FUNCTION_BLOCK FB_Line_Target EXTENDS FB_SFC_Cycle IMPLEMENTS ITF_FB_SFC_Cycle
VAR_INPUT
	valTankA				:	E_Pis_Name	;
	valTankB				:	E_Pis_Name	;
	valTankA_Pipe			:	E_Pis_Name	;
	valTankB_Pipe			:	E_Pis_Name	;
	valDrain				:	E_Pis_Name	;
	valCIP					:	E_Pis_Name	;
END_VAR
VAR_OUTPUT
END_VAR
VAR
	eReq				: E_Line_Target;
	eProcess			: E_Line_Target;
	eStatus				: E_Line_Target;
	
	fbPis				: FB_Piston;
	
	stPis_TankA				: REFERENCE TO ST_Piston;
	stPis_TankB				: REFERENCE TO ST_Piston;
	stPis_TankA_Pipe		: REFERENCE TO ST_Piston;
	stPis_TankB_Pipe		: REFERENCE TO ST_Piston;
	stPis_Drain				: REFERENCE TO ST_Piston;
	stPis_CIP				: REFERENCE TO ST_Piston;
	
	stPis_Outlet: ST_Piston;
	tonDrainTime: TON;
	rt_Req_Reset: R_TRIG;
END_VAR

act_GetReference();

act_Oper();
//IF NOT Init.x THEN
	act_Status();
//END_IF

tonDrainTime(PT:=T#1M, IN:=eStatus=E_Line_Target.eDrain AND eReq=E_Line_Target.eNone);
IF tonDrainTime.Q 
AND eReq=E_Line_Target.eNone
AND eProcess=E_Line_Target.eNone
THEN;
	eReq:=E_Line_Target.eClose;
END_IF

m_Request_Reset(memo:=rt_Req_Reset);//

ACTION _aCIP_active:
bStepDone:=FALSE;
IF TRUE 
AND eStatus=E_Line_Target.eCIP
THEN;
	bStepDone:=TRUE;
END_IF
END_ACTION

ACTION _aCIP_entry:
fbPis.m_SetByRecipe(stPis:=stPis_TankA, 			req:=E_Piston_Recipe_State.Release);
//fbPis.m_SetByRecipe(stPis:=stPis_TankA_Pipe, 		req:=E_Piston_Recipe_State.Release);		
fbPis.m_SetByRecipe(stPis:=stPis_TankB, 			req:=E_Piston_Recipe_State.Release);
//fbPis.m_SetByRecipe(stPis:=stPis_TankB_Pipe, 		req:=E_Piston_Recipe_State.Release);
fbPis.m_SetByRecipe(stPis:=stPis_Drain, 			req:=E_Piston_Recipe_State.Act);
fbPis.m_SetByRecipe(stPis:=stPis_CIP, 				req:=E_Piston_Recipe_State.Act);
END_ACTION

ACTION _aClose_active:
bStepDone:=FALSE;
IF TRUE 
AND eStatus=E_Line_Target.eClose
THEN;
	bStepDone:=TRUE;
END_IF
END_ACTION

ACTION _aClose_entry:
fbPis.m_SetByRecipe(stPis:=stPis_TankA, 			req:=E_Piston_Recipe_State.Release);
//fbPis.m_SetByRecipe(stPis:=stPis_TankA_Pipe, 		req:=E_Piston_Recipe_State.Release);		
fbPis.m_SetByRecipe(stPis:=stPis_TankB, 			req:=E_Piston_Recipe_State.Release);
//fbPis.m_SetByRecipe(stPis:=stPis_TankB_Pipe, 		req:=E_Piston_Recipe_State.Release);
fbPis.m_SetByRecipe(stPis:=stPis_Drain, 			req:=E_Piston_Recipe_State.Release);
fbPis.m_SetByRecipe(stPis:=stPis_CIP, 				req:=E_Piston_Recipe_State.Release);
END_ACTION

ACTION _aDone_entry:
eProcess:=E_Line_Target.eNone;
eReq:=E_Line_Target.eNone;
bRun:=FALSE;
bDone:=TRUE;
END_ACTION

ACTION _aDrain_active:
bStepDone:=FALSE;
IF TRUE 
AND eStatus=E_Line_Target.eDrain
THEN;
	bStepDone:=TRUE;
END_IF
END_ACTION

ACTION _aDrain_entry:
fbPis.m_SetByRecipe(stPis:=stPis_TankA, 			req:=E_Piston_Recipe_State.Release);	
//fbPis.m_SetByRecipe(stPis:=stPis_TankA_Pipe, 		req:=E_Piston_Recipe_State.Release);	
fbPis.m_SetByRecipe(stPis:=stPis_TankB, 			req:=E_Piston_Recipe_State.Release);
//fbPis.m_SetByRecipe(stPis:=stPis_TankB_Pipe, 		req:=E_Piston_Recipe_State.Release);
fbPis.m_SetByRecipe(stPis:=stPis_Drain, 			req:=E_Piston_Recipe_State.Act);
fbPis.m_SetByRecipe(stPis:=stPis_CIP, 				req:=E_Piston_Recipe_State.Release);
END_ACTION

ACTION _aInit_active:
SFCReset:=FALSE;
END_ACTION

ACTION _aInit_exit:
eProcess:=E_Line_Target.eNone;
eReq:=E_Line_Target.eNone;
END_ACTION

ACTION _aReady_active:
CASE eReq OF
	E_Line_Target.eClose:;
			IF TRUE THEN;
				eProcess:=E_Line_Target.eClose;
			END_IF

	E_Line_Target.eTank_A:;
			IF TRUE THEN;
				eProcess:=E_Line_Target.eTank_A;
			END_IF	
			
	E_Line_Target.eTank_B:;
			IF TRUE THEN;
				eProcess:=E_Line_Target.eTank_B;
			END_IF	
			
	E_Line_Target.eCIP:;
			IF TRUE THEN;
				eProcess:=E_Line_Target.eCIP;
			END_IF	

	E_Line_Target.eDrain:;
			IF TRUE THEN;
				eProcess:=E_Line_Target.eDrain;
			END_IF	
		
END_CASE
END_ACTION

ACTION _aReady_exit:
bRun:=TRUE;
bDone:=FALSE;
END_ACTION

ACTION _aTank_A_active:
bStepDone:=FALSE;
IF TRUE  
AND eStatus=E_Line_Target.eTank_A 
THEN;
	bStepDone:=TRUE;
END_IF
END_ACTION

ACTION _aTank_A_entry:
fbPis.m_SetByRecipe(stPis:=stPis_TankA, 			req:=E_Piston_Recipe_State.Act);	
fbPis.m_SetByRecipe(stPis:=stPis_TankA_Pipe, 		req:=E_Piston_Recipe_State.Release);	
fbPis.m_SetByRecipe(stPis:=stPis_TankB, 			req:=E_Piston_Recipe_State.Release);
//fbPis.m_SetByRecipe(stPis:=stPis_TankB_Pipe, 		req:=E_Piston_Recipe_State.Release);
fbPis.m_SetByRecipe(stPis:=stPis_Drain, 			req:=E_Piston_Recipe_State.Release);
fbPis.m_SetByRecipe(stPis:=stPis_CIP, 				req:=E_Piston_Recipe_State.Release);
END_ACTION

ACTION _aTank_B_active:
bStepDone:=FALSE;
IF TRUE 
AND eStatus=E_Line_Target.eTank_B
THEN;
	bStepDone:=TRUE;
END_IF
END_ACTION

ACTION _aTank_B_entry:
fbPis.m_SetByRecipe(stPis:=stPis_TankA, 			req:=E_Piston_Recipe_State.Release);	
//fbPis.m_SetByRecipe(stPis:=stPis_TankA_Pipe, 		req:=E_Piston_Recipe_State.Release);	
fbPis.m_SetByRecipe(stPis:=stPis_TankB, 			req:=E_Piston_Recipe_State.Act);
fbPis.m_SetByRecipe(stPis:=stPis_TankB_Pipe, 		req:=E_Piston_Recipe_State.Release);
fbPis.m_SetByRecipe(stPis:=stPis_Drain, 			req:=E_Piston_Recipe_State.Release);
fbPis.m_SetByRecipe(stPis:=stPis_CIP, 				req:=E_Piston_Recipe_State.Release);
END_ACTION

ACTION act_GetReference:
m_Set_SFCFlags_Reference();
//refElement REF= fbElement[eElementID];
//refState_Long REF= fbElement[eElementID].eState_Long;

stPis_TankA				REF= g_Piston.stPis[valTankA];
stPis_TankB				REF= g_Piston.stPis[valTankB];
stPis_TankA_Pipe		REF= g_Piston.stPis[valTankA_Pipe];
stPis_TankB_Pipe		REF= g_Piston.stPis[valTankB_Pipe];
stPis_Drain				REF= g_Piston.stPis[valDrain];
stPis_CIP				REF= g_Piston.stPis[valCIP];
END_ACTION

ACTION act_Oper:
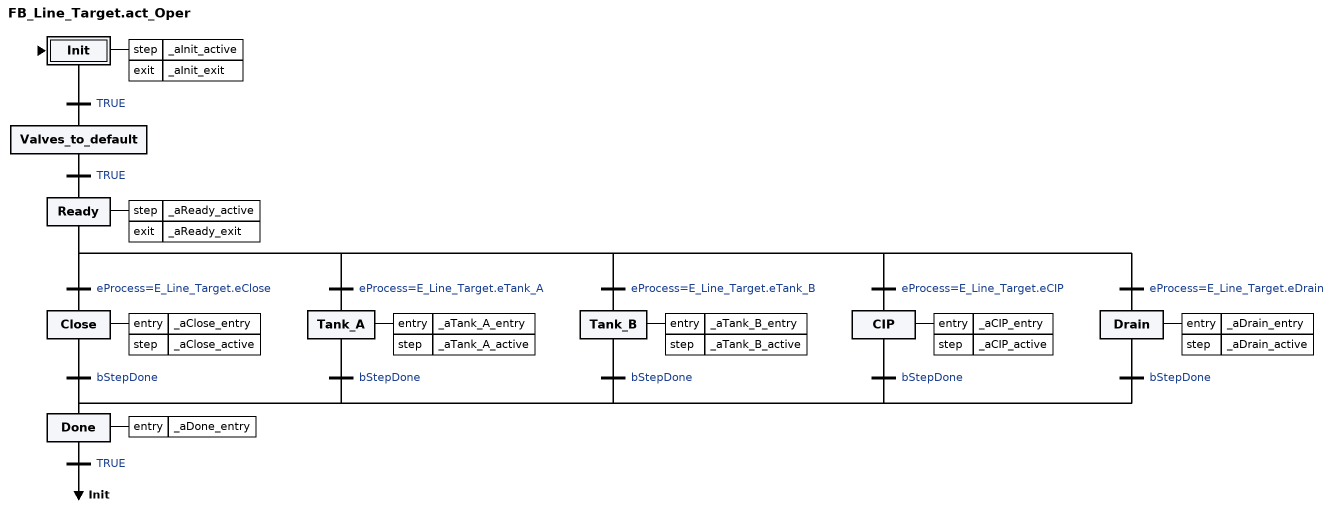
INITIAL_STEP Init:
    _aInit_active(N);  // step action
    _aInit_exit(P0);  // exit action
END_STEP
TRANSITION FROM Init TO Valves_to_default
    := TRUE;
END_TRANSITION
STEP Valves_to_default:
END_STEP
TRANSITION FROM Valves_to_default TO Ready
    := TRUE;
END_TRANSITION
STEP Ready:
    _aReady_active(N);  // step action
    _aReady_exit(P0);  // exit action
END_STEP
TRANSITION FROM Ready TO Close
    := eProcess=E_Line_Target.eClose;
END_TRANSITION
STEP Close:  // min time t#1s
    _aClose_entry(P1);  // entry action
    _aClose_active(N);  // step action
END_STEP
TRANSITION FROM Close TO Done
    := bStepDone;
END_TRANSITION
TRANSITION FROM Ready TO Tank_A
    := eProcess=E_Line_Target.eTank_A;
END_TRANSITION
STEP Tank_A:  // min time t#1s
    _aTank_A_entry(P1);  // entry action
    _aTank_A_active(N);  // step action
END_STEP
TRANSITION FROM Tank_A TO Done
    := bStepDone;
END_TRANSITION
TRANSITION FROM Ready TO Tank_B
    := eProcess=E_Line_Target.eTank_B;
END_TRANSITION
STEP Tank_B:  // min time t#1s
    _aTank_B_entry(P1);  // entry action
    _aTank_B_active(N);  // step action
END_STEP
TRANSITION FROM Tank_B TO Done
    := bStepDone;
END_TRANSITION
TRANSITION FROM Ready TO CIP
    := eProcess=E_Line_Target.eCIP;
END_TRANSITION
STEP CIP:  // min time t#1s
    _aCIP_entry(P1);  // entry action
    _aCIP_active(N);  // step action
END_STEP
TRANSITION FROM CIP TO Done
    := bStepDone;
END_TRANSITION
TRANSITION FROM Ready TO Drain
    := eProcess=E_Line_Target.eDrain;
END_TRANSITION
STEP Drain:  // min time t#1s
    _aDrain_entry(P1);  // entry action
    _aDrain_active(N);  // step action
END_STEP
TRANSITION FROM Drain TO Done
    := bStepDone;
END_TRANSITION
STEP Done:
    _aDone_entry(P1);  // entry action
END_STEP
TRANSITION FROM Done TO Init
    := TRUE;
END_TRANSITION
// branch label Branch0_act_Oper
END_ACTION

ACTION act_Status:
IF TRUE 
AND fbPis.m_CheckByRecipe(stPis:=stPis_TankA, 			req:=E_Piston_Recipe_State.Release)	
//AND fbPis.m_CheckByRecipe(stPis:=stPis_TankA_Pipe, 		req:=E_Piston_Recipe_State.Release)	
AND fbPis.m_CheckByRecipe(stPis:=stPis_TankB, 			req:=E_Piston_Recipe_State.Release)
//AND fbPis.m_CheckByRecipe(stPis:=stPis_TankB_Pipe, 		req:=E_Piston_Recipe_State.Release)
AND fbPis.m_CheckByRecipe(stPis:=stPis_Drain, 			req:=E_Piston_Recipe_State.Release)
AND fbPis.m_CheckByRecipe(stPis:=stPis_CIP, 			req:=E_Piston_Recipe_State.Release)
THEN;
	eStatus:=E_Line_Target.eClose;
ELSIF TRUE 
AND fbPis.m_CheckByRecipe(stPis:=stPis_TankA, 			req:=E_Piston_Recipe_State.Act)		
AND fbPis.m_CheckByRecipe(stPis:=stPis_TankA_Pipe, 		req:=E_Piston_Recipe_State.Release)	
AND fbPis.m_CheckByRecipe(stPis:=stPis_TankB, 			req:=E_Piston_Recipe_State.Release)
//AND fbPis.m_CheckByRecipe(stPis:=stPis_TankB_Pipe, 		req:=E_Piston_Recipe_State.Release)
AND fbPis.m_CheckByRecipe(stPis:=stPis_Drain, 			req:=E_Piston_Recipe_State.Release)
AND fbPis.m_CheckByRecipe(stPis:=stPis_CIP, 			req:=E_Piston_Recipe_State.Release)
THEN;
	eStatus:=E_Line_Target.eTank_A;
ELSIF TRUE 
AND fbPis.m_CheckByRecipe(stPis:=stPis_TankA, 			req:=E_Piston_Recipe_State.Release)		
//AND fbPis.m_CheckByRecipe(stPis:=stPis_TankA_Pipe, 		req:=E_Piston_Recipe_State.Release)	
AND fbPis.m_CheckByRecipe(stPis:=stPis_TankB, 			req:=E_Piston_Recipe_State.Act)
AND fbPis.m_CheckByRecipe(stPis:=stPis_TankB_Pipe, 		req:=E_Piston_Recipe_State.Release)
AND fbPis.m_CheckByRecipe(stPis:=stPis_Drain, 			req:=E_Piston_Recipe_State.Release)
AND fbPis.m_CheckByRecipe(stPis:=stPis_CIP, 			req:=E_Piston_Recipe_State.Release)
THEN;
	eStatus:=E_Line_Target.eTank_B;
ELSIF TRUE 
AND fbPis.m_CheckByRecipe(stPis:=stPis_TankA, 			req:=E_Piston_Recipe_State.Release)		
//AND fbPis.m_CheckByRecipe(stPis:=stPis_TankA_Pipe, 		req:=E_Piston_Recipe_State.Release)	
AND fbPis.m_CheckByRecipe(stPis:=stPis_TankB, 			req:=E_Piston_Recipe_State.Release)
//AND fbPis.m_CheckByRecipe(stPis:=stPis_TankB_Pipe, 		req:=E_Piston_Recipe_State.Release)
AND fbPis.m_CheckByRecipe(stPis:=stPis_Drain, 			req:=E_Piston_Recipe_State.Act)
AND fbPis.m_CheckByRecipe(stPis:=stPis_CIP, 			req:=E_Piston_Recipe_State.Act)
THEN;
	eStatus:=E_Line_Target.eCIP;
ELSIF TRUE 
AND fbPis.m_CheckByRecipe(stPis:=stPis_TankA, 			req:=E_Piston_Recipe_State.Release)		
//AND fbPis.m_CheckByRecipe(stPis:=stPis_TankA_Pipe, 		req:=E_Piston_Recipe_State.Release)	
AND fbPis.m_CheckByRecipe(stPis:=stPis_TankB, 			req:=E_Piston_Recipe_State.Release)
//AND fbPis.m_CheckByRecipe(stPis:=stPis_TankB_Pipe, 		req:=E_Piston_Recipe_State.Release)
AND fbPis.m_CheckByRecipe(stPis:=stPis_Drain, 			req:=E_Piston_Recipe_State.Act)
AND fbPis.m_CheckByRecipe(stPis:=stPis_CIP, 			req:=E_Piston_Recipe_State.Release)
THEN;
	eStatus:=E_Line_Target.eDrain;
ELSE;
	eStatus:=E_Line_Target.eNone;
END_IF
END_ACTION

METHOD m_CheckStatus : BOOL
VAR_INPUT
	eReqStatus		: E_Line_Target;
END_VAR
IF eStatus=eReqStatus 
AND eProcess=E_Line_Target.eNone
AND eReq=E_Line_Target.eNone
AND bReady
AND bDone
AND NOT bRun
THEN;
	m_CheckStatus:=TRUE;
END_IF
END_METHOD

METHOD m_Request_Reset : BOOL
VAR_IN_OUT
	memo: R_TRIG;
END_VAR
memo(CLK:=eReq=0);
IF TRUE 
AND memo.Q
THEN;
	SFCReset:=TRUE;
END_IF
END_METHOD

METHOD m_Run : BOOL
VAR_INPUT
	eReqProc			: E_Line_Target;
END_VAR
IF eProcess=E_Line_Target.eNone THEN;
	eProcess:=eReq:=eReqProc;
	bDone:=FALSE;
	m_Run:=TRUE;
END_IF
END_METHOD

METHOD m_Set_SFCFlags_Reference : BOOL
//Set reference to SFC flags

refSFC.SFCInit REF= SFCInit;
refSFC.SFCReset REF= SFCReset;
refSFC.SFCError REF= SFCError;
refSFC.SFCEnableLimit REF= SFCEnableLimit;
refSFC.SFCErrorStep REF= SFCErrorStep;
refSFC.SFCErrorPOU REF= SFCErrorPOU;
refSFC.SFCQuitError REF= SFCQuitError;
refSFC.SFCPause REF= SFCPause;
refSFC.SFCTrans REF= SFCTrans;
refSFC.SFCCurrentStep REF= SFCCurrentStep;
refSFC.SFCTip REF= SFCTip;
refSFC.SFCTipMode REF= SFCTipMode;

// Cycle handle for SFC
m_SFC_Handle();
END_METHOD

END_FUNCTION_BLOCK

(* stored: Version 1.1.0.1, ProductVersion 3.1.4024.15
   POU FB_Line_Target: Id {a73be08b-a059-412e-9240-f16489ac4962}, SpecialFunc None
   Folder Manage: Id {e5743553-9439-4305-9e84-949d6d5f1f58}
   Action _aCIP_active: Id {1c5f0b2c-a2c3-4aa0-90cb-5189c5a6156b}
   Action _aCIP_entry: Id {162310eb-2bb6-431e-b347-1831ed1ae816}
   Action _aClose_active: Id {4eee4bc2-b7ef-4e03-88f5-c6d6fb3b3622}
   Action _aClose_entry: Id {0e56069f-368f-4cd6-b1bd-6a8c8b618221}
   Action _aDone_entry: Id {ace91bfe-eb50-4697-9e26-19f420379f6a}
   Action _aDrain_active: Id {16bd941f-d65c-46b7-afee-66ba2e81eb6d}
   Action _aDrain_entry: Id {e3786de5-7c06-4103-8b0a-d372c40a7876}
   Action _aInit_active: Id {8a00560f-74f4-42ea-ad69-c17f7f4c4676}
   Action _aInit_exit: Id {699d0b5d-a3af-44d6-9603-9f23437535c9}
   Action _aReady_active: Id {9dae6a82-6750-4aef-88f6-30fbe0672b63}
   Action _aReady_exit: Id {991d30c6-bdb3-4d67-8d37-d97b5a4fe6b2}
   Action _aTank_A_active: Id {11e988fc-4330-4d0d-b9fd-24a06f163182}
   Action _aTank_A_entry: Id {2451655f-1f9c-46d1-bcc3-f92208ba93ea}
   Action _aTank_B_active: Id {1abd18c4-5659-4c67-8d8d-71c43176571d}
   Action _aTank_B_entry: Id {0e5f6a4c-494c-482b-8faf-2288a342d2b2}
   Action act_GetReference: Id {a3ab97cc-223f-4ca6-a0d8-38cc9345b8fd}
   Action act_Oper: Id {b85f536a-f031-4323-8005-3b43c10e0de6}
   Action act_Status: Id {8c31a424-7f78-49e2-b4ec-e3d2a2df1502}
   Method m_CheckStatus: Id {a95850ca-15b2-4e7e-a635-56b44d398318}
   Method m_Request_Reset: Id {95945eb0-2ad1-49de-8030-be298be214ee}
   Method m_Run: Id {4181f26e-983c-4e66-bf41-bf25464233de}
   Method m_Set_SFCFlags_Reference: Id {98131e4f-ae98-4828-8ba6-dcfb4bcb3c2f} *)
